{region 'Documentation'}
(*!
<summary>Check that IN is less than Maximum.</summary>
<description>

All checked operands and bounds must be finite; NaN or either infinity reports Error
during active evaluation.

Numeric diagnostics use the formatter's default six significant digits; rounding affects
the message only, not the comparison.

</description>
*)
{endregion}
FUNCTION_BLOCK AssertLessThan_Real EXTENDS AssertionBase
VAR_INPUT
    IN : REAL; //! Actual value checked or observed by this Assertion.
    Maximum : REAL; //! Exclusive upper bound; the actual value or count must be smaller.
END_VAR

SUPER^();

{region 'Documentation'}
(*!
<summary>Check that IN is less than Maximum.</summary>
*)
{endregion}
METHOD PROTECTED Assert
VAR
    Message : STRING(GVL_Constants.MessageLength);
    MaximumText : STRING(GVL_Constants.AssertionValueLength);
    ActualText : STRING(GVL_Constants.AssertionValueLength);
END_VAR
IF NOT EvaluationActive THEN
    RETURN;
END_IF;

IF Result = E_Result.Error THEN
    RETURN;
END_IF;

IF NOT Tc2_Utilities.RealIsFinite(x := IN) THEN
    Error(Message := 'Assertion error: IN must be finite.');
    RETURN;
END_IF;

IF NOT Tc2_Utilities.RealIsFinite(x := Maximum) THEN
    Error(Message := 'Assertion error: Maximum must be finite.');
    RETURN;
END_IF;

IF Result = E_Result.Failed THEN
    RETURN;
END_IF;

IF IN >= Maximum THEN
    MaximumText := CreateAssertionTextValue_Real(Value := Maximum);
    ActualText := CreateAssertionTextValue_Real(Value := IN);
    Message := CONCAT('Assertion failed: value is not less than maximum. Maximum = ',
        MaximumText);
    Message := CONCAT(Message, ', Actual = ');
    Message := CONCAT(Message, ActualText);
    Message := CONCAT(Message, '.');
    Fail(Message := Message);
    RETURN;
END_IF;

Pass();
END_METHOD

END_FUNCTION_BLOCK

(* stored: Version 1.1.0.1
   POU AssertLessThan_Real: Id {d20de2bd-0da4-4c54-9cf4-a86356f0b201}, SpecialFunc None
   Folder Internal: Id {176e54a0-c493-4ef8-ba0a-b44fbccfd063}
   Method Assert: Id {6f896d82-bb4b-434a-8d3d-7b0356b95a2c} *)
